// TIA Portal project "Plcs" (V21)

(* hardware
DEVICE "PLC_North"  S7-1500 station
   slot 0: "Rail_0"  Rack  6ES7 590-1***0-0AA0
   slot 1: "PLC_North"  CPU 1516-3 PN/DP  6ES7 516-3AN02-0AB0  V2.9
      slot 3: "CPU display_1"  6ES7591-1BA00-0AA0
      slot 32768: "PROFINET interface_1"  X1
         slot 32769: "Port_1"  X1 P1
         slot 32770: "Port_2"  X1 P2
      slot 33024: "PROFINET interface_2"  X2
         slot 33025: "Port_1"  X2 P1
      slot 33280: "DP interface_1"  X3
      slot 34817: "Virtual CP interface port_1"  Virtual CP interface port  Virtual CP interface port
DEVICE "PLC_South"  S7-1500 station
   slot 0: "Rail_0"  Rack  6ES7 590-1***0-0AA0
   slot 1: "PLC_South"  CPU 1516-3 PN/DP  6ES7 516-3AN02-0AB0  V2.9
      slot 3: "CPU display_1"  6ES7591-1BA00-0AA0
      slot 32768: "PROFINET interface_1"  X1
         slot 32769: "Port_1"  X1 P1
         slot 32770: "Port_2"  X1 P2
      slot 33024: "PROFINET interface_2"  X2
         slot 33025: "Port_1"  X2 P1
      slot 33280: "DP interface_1"  X3
      slot 34817: "Virtual CP interface port_1"  Virtual CP interface port  Virtual CP interface port
*)

// ===== PLC "PLC_North"  CPU 1516-3 PN/DP =====

VAR_GLOBAL   // PLC tag table "Counters"
   "Count_North" AT %MD0 : DInt;   // Starts counted on the north side
END_VAR

VAR_GLOBAL   // PLC tag table "IO"
   "Run_North" AT %I0.0 : Bool;   // Start the north station
   "Lamp_North" AT %Q0.0 : Bool;   // The north station runs
END_VAR

// folder: Area/Shared

TYPE "typeStatus"
   STRUCT
      running : Bool;   // Runs, north
      faults : Int;   // Faults counted on the north side
   END_STRUCT;
END_TYPE

// folder: Area/Data

DATA_BLOCK "StationData"   // DB1
{ S7_Optimized_Access := 'TRUE' }
VERSION : 0.1
// stored: InstanceOfName Station
"Station"
BEGIN
END_DATA_BLOCK

// folder: (top level)

ORGANIZATION_BLOCK "Main"   // OB1, SCL, ProgramCycle
TITLE = "Main Program Sweep (Cycle)"
{ S7_Optimized_Access := 'TRUE' }
VERSION : 0.1
   VAR_INPUT
      Initial_Call : Bool;   // Initial call of this OB
      Remanence : Bool;   // =True, if remanent data are available
   END_VAR
BEGIN

    "StationData"(run := "Run_North");
END_ORGANIZATION_BLOCK

// folder: Area/Line/Cell/Station

FUNCTION_BLOCK "Pump"   // FB1, SCL
TITLE = Pump of the north side
{ S7_Optimized_Access := 'TRUE' }
VERSION : 0.1
// One pump; the north PLC has a block of the same name with other text.
   VAR_INPUT
      run : Bool;   // Run the pump
   END_VAR
   VAR_OUTPUT
      status : "typeStatus";   // What the pump does
   END_VAR
BEGIN

    #status.running := #run;   // north
END_FUNCTION_BLOCK

FUNCTION_BLOCK "Station"   // FB2, SCL
TITLE = Station with 2 pumps
{ S7_Optimized_Access := 'TRUE' }
VERSION : 0.1
   VAR_INPUT
      run : Bool;   // Run the station
   END_VAR
   VAR
      pump1 : "Pump";   // Pump 1 of 2
      pump2 : "Pump";   // Pump 2 of 2
   END_VAR
BEGIN

    #pump1(run := #run);
    #pump2(run := #run);
END_FUNCTION_BLOCK

// ===== PLC "PLC_South"  CPU 1516-3 PN/DP =====

VAR_GLOBAL   // PLC tag table "Counters"
   "Count_South" AT %MD32 : DInt;   // Starts counted on the south side
END_VAR

VAR_GLOBAL   // PLC tag table "IO"
   "Run_South" AT %I8.0 : Bool;   // Start the south station
   "Lamp_South" AT %Q8.0 : Bool;   // The south station runs
END_VAR

// folder: Area/Shared

TYPE "typeStatus"
   STRUCT
      running : Bool;   // Runs, south
      faults : Int;   // Faults counted on the south side
   END_STRUCT;
END_TYPE

// folder: Area/Data

DATA_BLOCK "StationData"   // DB1
{ S7_Optimized_Access := 'TRUE' }
VERSION : 0.1
// stored: InstanceOfName Station
"Station"
BEGIN
END_DATA_BLOCK

// folder: (top level)

ORGANIZATION_BLOCK "Main"   // OB1, SCL, ProgramCycle
TITLE = "Main Program Sweep (Cycle)"
{ S7_Optimized_Access := 'TRUE' }
VERSION : 0.1
   VAR_INPUT
      Initial_Call : Bool;   // Initial call of this OB
      Remanence : Bool;   // =True, if remanent data are available
   END_VAR
BEGIN

    "StationData"(run := "Run_South");
END_ORGANIZATION_BLOCK

// folder: Area/Line/Cell/Station

FUNCTION_BLOCK "Pump"   // FB1, SCL
TITLE = Pump of the south side
{ S7_Optimized_Access := 'TRUE' }
VERSION : 0.1
// One pump; the south PLC has a block of the same name with other text.
   VAR_INPUT
      run : Bool;   // Run the pump
   END_VAR
   VAR_OUTPUT
      status : "typeStatus";   // What the pump does
   END_VAR
BEGIN

    #status.running := #run;   // south
END_FUNCTION_BLOCK

FUNCTION_BLOCK "Station"   // FB2, SCL
TITLE = Station with 3 pumps
{ S7_Optimized_Access := 'TRUE' }
VERSION : 0.1
   VAR_INPUT
      run : Bool;   // Run the station
   END_VAR
   VAR
      pump1 : "Pump";   // Pump 1 of 3
      pump2 : "Pump";   // Pump 2 of 3
      pump3 : "Pump";   // Pump 3 of 3
   END_VAR
BEGIN

    #pump1(run := #run);
    #pump2(run := #run);
    #pump3(run := #run);
END_FUNCTION_BLOCK